(* IEC 61131-3 sources: rusty/tests/lit/cfc/validation/unresolved_reference, 1 file *)

(* ---- main.st ---- *)
// Sources and sinks naming undeclared variables, also nested in a global access and in an array
// literal, with and without parentheses. Each unresolved reference is reported at its sink block;
// a source has no execution order and is located at the sink it feeds.
// CHECK: {{.*}}unresolved_reference.cfc.unresolved_reference:1: error[E048]: Could not resolve reference to foo
// CHECK: {{.*}}unresolved_reference.cfc.unresolved_reference:1: error[E048]: Could not resolve reference to asd
// CHECK: {{.*}}unresolved_reference.cfc.unresolved_reference:2: error[E048]: Could not resolve reference to global
// CHECK: {{.*}}unresolved_reference.cfc.unresolved_reference:3: error[E048]: Could not resolve reference to element
// CHECK: {{.*}}unresolved_reference.cfc.unresolved_reference:4: error[E048]: Could not resolve reference to parenGlobal
// CHECK: {{.*}}unresolved_reference.cfc.unresolved_reference:5: error[E048]: Could not resolve reference to parenElement
// CHECK: error: Compilation aborted due to critical errors
FUNCTION main : DINT
END_FUNCTION
